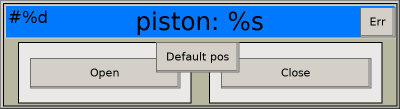
VISUALIZATION vis_Piston_Control1_Compact  // 400x109
VAR_IN_OUT
	stPis: ST_Piston;
END_VAR
    Rectangle (0,0 400x109)
    Rectangle (3,3 394x103), colour toggle: NOT stPis.b_Enable
    Rectangle (18,42 173x61), colour toggle: stPis.st_Open
    Rectangle (209,42 173x61), colour toggle: stPis.st_Close
    Button (30,58 150x30), "Open", colour toggle: stPis.req_Open, input disabled if: stPis.b_DeactivateMan OR NOT stPis.b_InterLock_Open
        toggle stPis.req_OpenMan
    Button (221,58 150x30), "Close", colour toggle: stPis.req_Close, input disabled if: stPis.b_DeactivateMan OR NOT stPis.b_InterLock_Close
        toggle stPis.req_CloseMan
    Button (156,42 83x30), "Default pos", colour toggle: stPis.req_DefaultPos, input disabled if: stPis.b_DeactivateMan
        toggle stPis.req_DefaultPos
    Textfield (5,5 390x33), "piston: %s", text variable: stPis.sName
    Textfield (5,7 42x21), "#%d", text variable: stPis.iPisNum
    Button (360,7 35x30), "Err", colour toggle: stPis.b_Error
        toggle stPis.b_Resume
END_VISUALIZATION

(* stored: Version 1.1.0.1, ProductVersion 3.1.4024.12
   Visu vis_Piston_Control1_Compact: Id {e0c313ee-4f7e-40c8-bbf0-f3c25540c374} *)
